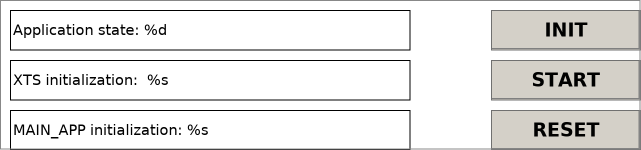
VISUALIZATION T_MAIN_APP  // 641x150
VAR_IN_OUT
	DataIn    : ST_MAIN_VIS;
  DataOut   : ST_VIS_MAIN;
END_VAR
    Rectangle (10,10 400x40), "Application state: %d", text variable: DataIn.nStateApplication
    Rectangle (10,60 400x40), "XTS initialization: %s", text variable: DataIn.sInitXts, colour toggle: (DataIn.eInitXts = E_PROGRESS.PROGRESS_DONE)
    Rectangle (10,110 400x40), "MAIN_APP initialization: %s", text variable: DataIn.sInitApplication, colour toggle: (DataIn.eInitApplication = E_PROGRESS.PROGRESS_DONE)
    Button (491,10 150x40), "INIT"
        toggle DataOut.Init
    Button (491,60 150x40), "START"
        tap DataOut.Start
    Button (491,110 150x40), "RESET"
        tap DataOut.Reset
END_VISUALIZATION

(* stored: Version 1.1.0.1, ProductVersion 3.1.4026.20
   Visu T_MAIN_APP: Id {92f746a9-8bb1-41ea-942c-20b90b4af519} *)
